(* IEC 61131-3 sources: llm-plc-st-eval/data/processed_definitivo/qwen2.5-coder_14b/B1/zero_shot, 3 files *)

(* ---- ejec_1.st ---- *)
FUNCTION_BLOCK FB_Motor
VAR_INPUT
    btnMarcha : BOOL;  // Botón de marcha
    btnParo : BOOL;    // Botón de paro
    btnEmerg : BOOL;   // Botón de paro de emergencia
END_VAR

VAR_OUTPUT
    motorOn : BOOL;    // Estado del motor (encendido/apagado)
END_VAR

VAR
    emergenciaActiva : BOOL := FALSE;  // Bandera para indicar si hay una parada de emergencia
END_VAR

// Programa principal
IF btnEmerg THEN
    // Si se activa el botón de emergencia, detener el motor y activar la bandera de emergencia
    motorOn := FALSE;
    emergenciaActiva := TRUE;
ELSIF emergenciaActiva THEN
    // Si hay una parada de emergencia activa, mantener el motor apagado
    motorOn := FALSE;
ELSIF btnParo THEN
    // Si se presiona el botón de paro, detener el motor
    motorOn := FALSE;
ELSIF btnMarcha THEN
    // Si se presiona el botón de marcha, encender el motor
    motorOn := TRUE;
END_IF;

(* ---- ejec_2.st ---- *)
FUNCTION_BLOCK FB_Motor
VAR_INPUT
    btnMarcha : BOOL;  // Botón de marcha
    btnParo : BOOL;    // Botón de paro
    btnEmerg : BOOL;   // Botón de paro de emergencia
END_VAR

VAR_OUTPUT
    motorOn : BOOL;    // Estado del motor (encendido/apagado)
END_VAR

VAR
    emergenciaActiva : BOOL := FALSE;  // Bandera para indicar si hay una emergencia activa
END_VAR

// Programa principal
IF btnEmerg THEN
    // Si se activa el botón de emergencia
    emergenciaActiva := TRUE;
    motorOn := FALSE;  // Apaga el motor
ELSEIF emergenciaActiva THEN
    // Si hay una emergencia activa, no se permite el arranque del motor
    motorOn := FALSE;
ELSEIF btnParo THEN
    // Si se presiona el botón de paro
    motorOn := FALSE;  // Apaga el motor
ELSEIF btnMarcha THEN
    // Si se presiona el botón de marcha
    motorOn := TRUE;   // Enciende el motor
END_IF;

(* ---- ejec_3.st ---- *)
FUNCTION_BLOCK FB_Motor
VAR_INPUT
    btnMarcha : BOOL;  // Botón de marcha
    btnParo : BOOL;    // Botón de paro
    btnEmerg : BOOL;   // Botón de paro de emergencia
END_VAR

VAR_OUTPUT
    motorOn : BOOL;    // Estado del motor (encendido/apagado)
END_VAR

VAR
    emergenciaActiva : BOOL := FALSE;  // Bandera para indicar si hay una parada de emergencia
END_VAR

// Programa principal
IF btnEmerg THEN
    // Si se detecta una parada de emergencia
    emergenciaActiva := TRUE;
    motorOn := FALSE;  // Apaga el motor
ELSEIF emergenciaActiva THEN
    // Si hay una parada de emergencia activa, no se permite el arranque
    motorOn := FALSE;
ELSEIF btnParo THEN
    // Si se presiona el botón de paro
    motorOn := FALSE;  // Apaga el motor
ELSEIF btnMarcha THEN
    // Si se presiona el botón de marcha
    motorOn := TRUE;   // Enciende el motor
END_IF
